PROGRAM main
  VAR
    B1 AT %IX0.0  : BOOL; (* sensor de piezas *)
    S1 AT %IX0.1  : BOOL; (* RESET *)
    KM1 AT %QX0.0 : BOOL; (* motor de la cinta *)
    H1 AT %QX0.1  : BOOL; (* caja llena *)
    PIEZAS        : CTU;
    LLENA         : BOOL;
    CUENTA        : INT; (* piezas en la caja *)
  END_VAR
  VAR  (* added by the conversion: wires and edge detectors of the diagram *)
    _NOT7_OUT : BOOL;
  END_VAR

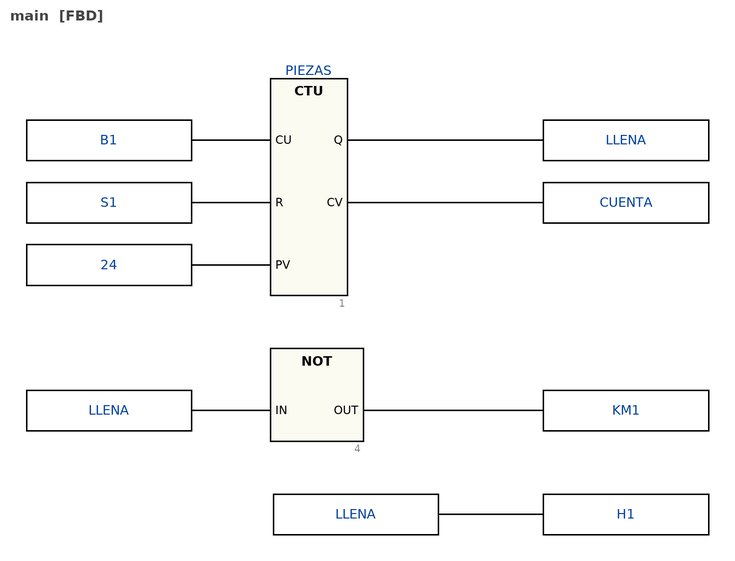
(* FBD diagram, written out as Structured Text *)
PIEZAS(CU := B1, R := S1, PV := 24);
LLENA := PIEZAS.Q;
CUENTA := PIEZAS.CV;
_NOT7_OUT := NOT LLENA;
KM1 := _NOT7_OUT;
H1 := LLENA;
END_PROGRAM
